(****************************************************************************************************<br>
© Syntegon Group.<br>
All rights reserved, also regarding any disposal, exploitation, reproduction, editing, distribution,<br>
as well as in the event of applications for industrial property rights.<br>
*****************************************************************************************************<br>
DESCRIPTION:<br>
Passes the effective pose, origin shift and zones on to the component's Syn_Visu FB; for m_PassOn of the<br>
derived FB, which knows where the visualisation keeps its zone count.<br>
****************************************************************************************************)
METHOD PROTECTED m_PassOnBody : BOOL
VAR_IN_OUT
	vio_Visu							: SynVisu._FB_VisuBodyComponent;	// the component's Syn_Visu FB
END_VAR
VAR_INPUT
	vi_un_VisuZoneCount					: UINT;	// [-] zones the visualisation has now, its stConfig.nZoneCount
END_VAR
m_PassOnBody := TRUE;
vio_Visu.m_SetPose(vi_Pose := vo_Config.stActive.stPose);
vio_Visu.m_SetOriginShift(vi_lr_X := vo_Config.stActive.stOriginShift.fX, vi_lr_Y := vo_Config.stActive.stOriginShift.fY,
	vi_lr_Z := vo_Config.stActive.stOriginShift.fZ);
m_PassOnZones(vio_Visu := vio_Visu, vio_aZones := vo_Config.stActive.aZones, vi_un_Count := vo_Config.stActive.nZoneCount,
	vi_un_VisuCount := vi_un_VisuZoneCount);
END_METHOD

(****************************************************************************************************<br>
© Syntegon Group.<br>
All rights reserved, also regarding any disposal, exploitation, reproduction, editing, distribution,<br>
as well as in the event of applications for industrial property rights.<br>
*****************************************************************************************************<br>
DESCRIPTION:<br>
Effective pose (MCS), for the application's logic.<br>
****************************************************************************************************)
METHOD m_Pose : SynVisu.ST_VisuPose
m_Pose := vo_Config.stActive.stPose;
END_METHOD

END_FUNCTION_BLOCK

// ---- POUs/_FB_ConfigCartesian.TcPOU
(****************************************************************************************************<br>
© Syntegon Group.<br>
All rights reserved, also regarding any disposal, exploitation, reproduction, editing, distribution,<br>
as well as in the event of applications for industrial property rights.<br>
*****************************************************************************************************<br>
DESCRIPTION:<br>
Parameter set of one Cartesian robot (ADR 0017): its pose, origin shift, zones, gripper fingers, limit area and<br>
TCP limit area, written by the configurator, taken over when the application allows it.<br>
Typical cycle:<br>
  fb_CartParam.m_Register(vio_Manifest := GVL_Config.stManifest, vi_udn_Id := fb_Cart.m_Id());<br>
  fb_CartParam.m_Cycle(vio_Default := CartDefault, vio_Set := CartSet, vi_b_ApplyAllowed := b_Stopped);<br>
  fb_Cart.m_Configure(vi_lr_XMin := 0, ...);<br>
  fb_CartParam.m_PassOn(vio_Visu := fb_Cart);<br>
The application's logic takes its zones and limit areas from m_Active, not from its own constants.<br>
*****************************************************************************************************<br>
OUTPUT VALUES:<br>
vo_Config is the contract structure the gateway reads and writes at the path in the config manifest.<br>
*****************************************************************************************************<br>
VERSION         ¦ DATE       ¦ NAME      ¦ CHANGE<br>
Syn_Config 1.1.0 ¦ 2026-11-10 ¦ J.Willner ¦ New<br>
Syn_Config 2.0.0 ¦ 2026-11-11 ¦ J.Willner ¦ Gripper fingers with their offsets, m_Invalid (ADR 0018)<br>
Syn_Config 2.3.0 ¦ 2026-11-14 ¦ J.Willner ¦ m_Cycle through m_HandleStaging; m_PassOn passes the pose on<br>
****************************************************************************************************)
FUNCTION_BLOCK _FB_ConfigCartesian EXTENDS _FB_ConfigComponent
VAR_OUTPUT
	vo_Config							: ST_ConfigCartesian;	// contract structure of the gateway
END_VAR

(****************************************************************************************************<br>
© Syntegon Group.<br>
All rights reserved, also regarding any disposal, exploitation, reproduction, editing, distribution,<br>
as well as in the event of applications for industrial property rights.<br>
*****************************************************************************************************<br>
DESCRIPTION:<br>
All effective values (zones, limit areas, ...), for the application's own logic.<br>
****************************************************************************************************)
METHOD m_Active : ST_ConfigCartesianParam
m_Active := vo_Config.stActive;
END_METHOD

(****************************************************************************************************<br>
© Syntegon Group.<br>
All rights reserved, also regarding any disposal, exploitation, reproduction, editing, distribution,<br>
as well as in the event of applications for industrial property rights.<br>
*****************************************************************************************************<br>
DESCRIPTION:<br>
A Cartesian robot.<br>
****************************************************************************************************)
METHOD PROTECTED m_ComponentType : SynVisu.E_VisuComponentType
m_ComponentType := SynVisu.E_VisuComponentType.CARTESIAN;
END_METHOD

(****************************************************************************************************<br>
© Syntegon Group.<br>
All rights reserved, also regarding any disposal, exploitation, reproduction, editing, distribution,<br>
as well as in the event of applications for industrial property rights.<br>
*****************************************************************************************************<br>
DESCRIPTION:<br>
Every cycle: handles a staged set or a reset (a set only while vi_b_ApplyAllowed), keeps the active set in<br>
vio_Set and gives the effective values in vo_Config.stActive: the active set while one is valid, else the<br>
program values vio_Default.<br>
*****************************************************************************************************<br>
OUTPUT VALUES:<br>
TRUE in the cycle a set was taken over or reset.<br>
****************************************************************************************************)
METHOD m_Cycle : BOOL
VAR_IN_OUT CONSTANT
	vio_Default							: ST_ConfigCartesianParam;	// the application's program values
END_VAR
VAR_IN_OUT
	vio_Set								: ST_ConfigCartesianSet;	// the application's VAR PERSISTENT active set
END_VAR
VAR_INPUT
	vi_b_ApplyAllowed					: BOOL;	// [-] a staged set may be taken over now, e.g. while the machine stands
END_VAR
VAR
	b_TempTakeOver						: BOOL;	// the staged set was taken over: copy it
END_VAR
m_Cycle := m_HandleStaging(vio_Staging := vo_Config.stStaging, vio_Status := vo_Config.stStatus, vio_b_Valid := vio_Set.bValid,
	vio_udn_Version := vio_Set.nVersion, vio_udn_LastVersion := vio_Set.nLastVersion, vi_b_ApplyAllowed := vi_b_ApplyAllowed,
	vo_b_TakeOver => b_TempTakeOver);
IF b_TempTakeOver THEN
	vio_Set.stParam := vo_Config.stStaged;
END_IF


(****************************************************************************************************
EFFECTIVE VALUES
****************************************************************************************************)
IF vio_Set.bValid THEN
	vo_Config.stActive := vio_Set.stParam;
ELSE
	vo_Config.stActive := vio_Default;
END_IF
END_METHOD

(****************************************************************************************************<br>
© Syntegon Group.<br>
All rights reserved, also regarding any disposal, exploitation, reproduction, editing, distribution,<br>
as well as in the event of applications for industrial property rights.<br>
*****************************************************************************************************<br>
DESCRIPTION:<br>
Why a staged set cannot be taken over; '' when it can: more zones or fingers than the lists hold, a zone on no<br>
conveyor (id 0), or a finger without a diameter or height.<br>
****************************************************************************************************)
METHOD PROTECTED m_InvalidStaged : STRING(80)
m_InvalidStaged := m_InvalidZones(vio_aZones := vo_Config.stStaged.aZones, vi_un_Count := vo_Config.stStaged.nZoneCount);
IF m_InvalidStaged = '' THEN
	m_InvalidStaged := m_InvalidFingers(vio_aFingers := vo_Config.stStaged.aFingers, vi_un_Count := vo_Config.stStaged.nFingerCount);
END_IF
END_METHOD

(****************************************************************************************************<br>
© Syntegon Group.<br>
All rights reserved, also regarding any disposal, exploitation, reproduction, editing, distribution,<br>
as well as in the event of applications for industrial property rights.<br>
*****************************************************************************************************<br>
DESCRIPTION:<br>
Passes the effective pose, origin shift, limit areas, zones and fingers on to the robot's Syn_Visu FB, so the<br>
visualisation shows what the machine uses; the strokes and rail height (hardware) stay with the application's<br>
m_Configure call. Call it after m_Cycle, every cycle; Syn_Visu's config version only changes when a value does.<br>
****************************************************************************************************)
METHOD m_PassOn : BOOL
VAR_IN_OUT
	vio_Visu							: SynVisu._FB_VisuCartesian;	// the robot's Syn_Visu FB
END_VAR
m_PassOn := TRUE;
vio_Visu.m_SetPose(vi_Pose := vo_Config.stActive.stPose);
vio_Visu.m_SetOriginShift(vi_lr_X := vo_Config.stActive.stOriginShift.fX, vi_lr_Y := vo_Config.stActive.stOriginShift.fY,
	vi_lr_Z := vo_Config.stActive.stOriginShift.fZ);
m_PassOnLimitAreas(vio_Visu := vio_Visu, vio_LimitArea := vo_Config.stActive.stLimitArea,
	vio_TcpLimitArea := vo_Config.stActive.stTcpLimitArea);
m_PassOnZones(vio_Visu := vio_Visu, vio_aZones := vo_Config.stActive.aZones, vi_un_Count := vo_Config.stActive.nZoneCount,
	vi_un_VisuCount := vio_Visu.vo_Visu.stConfig.nZoneCount);
m_PassOnFingers(vio_Visu := vio_Visu, vio_aFingers := vo_Config.stActive.aFingers,
	vi_un_Count := vo_Config.stActive.nFingerCount, vi_un_VisuCount := vio_Visu.vo_Visu.stConfig.nFingerCount);
END_METHOD

(****************************************************************************************************<br>
© Syntegon Group.<br>
All rights reserved, also regarding any disposal, exploitation, reproduction, editing, distribution,<br>
as well as in the event of applications for industrial property rights.<br>
*****************************************************************************************************<br>
DESCRIPTION:<br>
Effective pose of the axis origin (MCS), for the application's logic.<br>
****************************************************************************************************)
METHOD m_Pose : SynVisu.ST_VisuPose
m_Pose := vo_Config.stActive.stPose;
END_METHOD

END_FUNCTION_BLOCK

// ---- POUs/_FB_ConfigConveyor.TcPOU
(****************************************************************************************************<br>
© Syntegon Group.<br>
All rights reserved, also regarding any disposal, exploitation, reproduction, editing, distribution,<br>
as well as in the event of applications for industrial property rights.<br>
*****************************************************************************************************<br>
DESCRIPTION:<br>
Parameter set of one conveyor (ADR 0017): its pose, origin shift and product types, written by the configurator,<br>
taken over when the application allows it. Typical cycle, before the Syn_Visu calls of the conveyor:<br>
  fb_InfeedParam.m_Register(vio_Manifest := GVL_Config.stManifest, vi_udn_Id := fb_Infeed.m_Id());<br>
  fb_InfeedParam.m_Cycle(vio_Default := InfeedDefault, vio_Set := InfeedSet, vi_b_ApplyAllowed := b_Stopped);<br>
  fb_Infeed.m_Configure(vi_lr_Length := 3000, vi_lr_Width := 400);<br>
  fb_InfeedParam.m_PassOn(vio_Visu := fb_Infeed);<br>
InfeedSet is the application's VAR PERSISTENT ST_ConfigConveyorSet; InfeedDefault its program values.<br>
*****************************************************************************************************<br>
OUTPUT VALUES:<br>
vo_Config is the contract structure the gateway reads and writes at the path in the config manifest.<br>
*****************************************************************************************************<br>
VERSION         ¦ DATE       ¦ NAME      ¦ CHANGE<br>
Syn_Config 1.0.0 ¦ 2026-11-10 ¦ J.Willner ¦ First version<br>
Syn_Config 2.3.0 ¦ 2026-11-14 ¦ J.Willner ¦ m_Cycle through m_HandleStaging; m_PassOn passes the pose on<br>
****************************************************************************************************)
FUNCTION_BLOCK _FB_ConfigConveyor EXTENDS _FB_ConfigComponent
VAR_OUTPUT
	vo_Config							: ST_ConfigConveyor;	// contract structure of the gateway
END_VAR

(****************************************************************************************************<br>
© Syntegon Group.<br>
All rights reserved, also regarding any disposal, exploitation, reproduction, editing, distribution,<br>
as well as in the event of applications for industrial property rights.<br>
*****************************************************************************************************<br>
DESCRIPTION:<br>
All effective values (origin shift, product types, ...), for the application's own logic.<br>
****************************************************************************************************)
METHOD m_Active : ST_ConfigConveyorParam
m_Active := vo_Config.stActive;
END_METHOD

(****************************************************************************************************<br>
© Syntegon Group.<br>
All rights reserved, also regarding any disposal, exploitation, reproduction, editing, distribution,<br>
as well as in the event of applications for industrial property rights.<br>
*****************************************************************************************************<br>
DESCRIPTION:<br>
A conveyor.<br>
****************************************************************************************************)
METHOD PROTECTED m_ComponentType : SynVisu.E_VisuComponentType
m_ComponentType := SynVisu.E_VisuComponentType.CONVEYOR;
END_METHOD

(****************************************************************************************************<br>
© Syntegon Group.<br>
All rights reserved, also regarding any disposal, exploitation, reproduction, editing, distribution,<br>
as well as in the event of applications for industrial property rights.<br>
*****************************************************************************************************<br>
DESCRIPTION:<br>
Every cycle: handles a staged set or a reset (a set only while vi_b_ApplyAllowed), keeps the active set in<br>
vio_Set and gives the effective values in vo_Config.stActive: the active set while one is valid, else the<br>
program values vio_Default.<br>
*****************************************************************************************************<br>
OUTPUT VALUES:<br>
TRUE in the cycle a set was taken over or reset.<br>
****************************************************************************************************)
METHOD m_Cycle : BOOL
VAR_IN_OUT CONSTANT
	vio_Default							: ST_ConfigConveyorParam;	// the application's program values
END_VAR
VAR_IN_OUT
	vio_Set								: ST_ConfigConveyorSet;	// the application's VAR PERSISTENT active set
END_VAR
VAR_INPUT
	vi_b_ApplyAllowed					: BOOL;	// [-] a staged set may be taken over now, e.g. while the machine stands
END_VAR
VAR
	b_TempTakeOver						: BOOL;	// the staged set was taken over: copy it
END_VAR
m_Cycle := m_HandleStaging(vio_Staging := vo_Config.stStaging, vio_Status := vo_Config.stStatus, vio_b_Valid := vio_Set.bValid,
	vio_udn_Version := vio_Set.nVersion, vio_udn_LastVersion := vio_Set.nLastVersion, vi_b_ApplyAllowed := vi_b_ApplyAllowed,
	vo_b_TakeOver => b_TempTakeOver);
IF b_TempTakeOver THEN
	vio_Set.stParam := vo_Config.stStaged;
END_IF


(****************************************************************************************************
EFFECTIVE VALUES
****************************************************************************************************)
IF vio_Set.bValid THEN
	vo_Config.stActive := vio_Set.stParam;
ELSE
	vo_Config.stActive := vio_Default;
END_IF
END_METHOD

(****************************************************************************************************<br>
© Syntegon Group.<br>
All rights reserved, also regarding any disposal, exploitation, reproduction, editing, distribution,<br>
as well as in the event of applications for industrial property rights.<br>
*****************************************************************************************************<br>
DESCRIPTION:<br>
Why a staged set cannot be taken over; '' when it can: more product types than the list holds, a product type<br>
without a number or a number used twice.<br>
****************************************************************************************************)
METHOD PROTECTED m_InvalidStaged : STRING(80)
VAR
	un_TempIndex						: UINT;
	un_TempOther						: UINT;
END_VAR
m_InvalidStaged := '';
IF vo_Config.stStaged.nProductTypeCount > SynVisu.VISU_GlobalConst_Param.VISU_un_MAX_PRODUCT_TYPES THEN
	m_InvalidStaged := CONCAT('More than ', CONCAT(UINT_TO_STRING(SynVisu.VISU_GlobalConst_Param.VISU_un_MAX_PRODUCT_TYPES), ' product types'));
	RETURN;
END_IF
un_TempIndex := 0;
WHILE un_TempIndex < vo_Config.stStaged.nProductTypeCount DO
	IF vo_Config.stStaged.aProductTypes[un_TempIndex].nId = 0 THEN
		m_InvalidStaged := 'A product type without a number';
		RETURN;
	END_IF
	un_TempOther := 0;
	WHILE un_TempOther < un_TempIndex DO
		IF vo_Config.stStaged.aProductTypes[un_TempOther].nId = vo_Config.stStaged.aProductTypes[un_TempIndex].nId THEN
			m_InvalidStaged := CONCAT('Product type ',
				CONCAT(UDINT_TO_STRING(vo_Config.stStaged.aProductTypes[un_TempIndex].nId), ' is defined twice'));
			RETURN;
		END_IF
		un_TempOther := un_TempOther + 1;
	END_WHILE
	un_TempIndex := un_TempIndex + 1;
END_WHILE
END_METHOD

(****************************************************************************************************<br>
© Syntegon Group.<br>
All rights reserved, also regarding any disposal, exploitation, reproduction, editing, distribution,<br>
as well as in the event of applications for industrial property rights.<br>
*****************************************************************************************************<br>
DESCRIPTION:<br>
Passes the effective pose, origin shift and product types on to the conveyor's Syn_Visu FB, so the<br>
visualisation shows what the machine uses; the belt's length and width (hardware) stay with the application's<br>
m_Configure call. Call it after m_Cycle, every cycle; Syn_Visu's config version only changes when a value does.<br>
*****************************************************************************************************<br>
LIMITS:<br>
Syn_Visu cannot remove a product type: one the set no longer has stays in the visualisation until the<br>
application restarts (the configurator warns of the difference).<br>
****************************************************************************************************)
METHOD m_PassOn : BOOL
VAR_IN_OUT
	vio_Visu							: SynVisu._FB_VisuConveyor;	// the conveyor's Syn_Visu FB
END_VAR
VAR
	un_TempIndex						: UINT;
END_VAR
m_PassOn := TRUE;
vio_Visu.m_SetPose(vi_Pose := vo_Config.stActive.stPose);
vio_Visu.m_SetOriginShift(vi_lr_X := vo_Config.stActive.stOriginShift.fX, vi_lr_Y := vo_Config.stActive.stOriginShift.fY,
	vi_lr_Z := vo_Config.stActive.stOriginShift.fZ);
un_TempIndex := 0;
WHILE un_TempIndex < vo_Config.stActive.nProductTypeCount
	AND un_TempIndex < SynVisu.VISU_GlobalConst_Param.VISU_un_MAX_PRODUCT_TYPES
DO
	vio_Visu.m_SetProductType(vi_udn_Id := vo_Config.stActive.aProductTypes[un_TempIndex].nId,
		vi_lr_Length := vo_Config.stActive.aProductTypes[un_TempIndex].fLength,
		vi_lr_Width := vo_Config.stActive.aProductTypes[un_TempIndex].fWidth,
		vi_lr_Height := vo_Config.stActive.aProductTypes[un_TempIndex].fHeight,
		vi_e_Shape := vo_Config.stActive.aProductTypes[un_TempIndex].eShape,
		vi_lr_CornerRadius := vo_Config.stActive.aProductTypes[un_TempIndex].fCornerRadius);
	un_TempIndex := un_TempIndex + 1;
END_WHILE
END_METHOD

(****************************************************************************************************<br>
© Syntegon Group.<br>
All rights reserved, also regarding any disposal, exploitation, reproduction, editing, distribution,<br>
as well as in the event of applications for industrial property rights.<br>
*****************************************************************************************************<br>
DESCRIPTION:<br>
Effective pose of the belt start (MCS), for the application's logic.<br>
****************************************************************************************************)
METHOD m_Pose : SynVisu.ST_VisuPose
m_Pose := vo_Config.stActive.stPose;
END_METHOD

END_FUNCTION_BLOCK

// ---- POUs/_FB_ConfigDelta.TcPOU
(****************************************************************************************************<br>
© Syntegon Group.<br>
All rights reserved, also regarding any disposal, exploitation, reproduction, editing, distribution,<br>
as well as in the event of applications for industrial property rights.<br>
*****************************************************************************************************<br>
DESCRIPTION:<br>
Parameter set of one Delta robot (ADR 0017): its pose, origin shift, zones, gripper fingers, working area,<br>
limit area and TCP limit area, written by the configurator, taken over when the application allows it.<br>
Typical cycle:<br>
  fb_Delta1Param.m_Register(vio_Manifest := GVL_Config.stManifest, vi_udn_Id := fb_Delta1.m_Id());<br>
  fb_Delta1Param.m_Cycle(vio_Default := Delta1Default, vio_Set := Delta1Set, vi_b_ApplyAllowed := b_Stopped);<br>
  fb_Delta1.m_Configure(vi_lr_BaseRadius := 200, ...);<br>
  fb_Delta1Param.m_PassOn(vio_Visu := fb_Delta1);<br>
The application's pick logic takes its zones from m_Zone / m_Active, not from its own constants.<br>
*****************************************************************************************************<br>
OUTPUT VALUES:<br>
vo_Config is the contract structure the gateway reads and writes at the path in the config manifest.<br>
*****************************************************************************************************<br>
VERSION         ¦ DATE       ¦ NAME      ¦ CHANGE<br>
Syn_Config 1.0.0 ¦ 2026-11-10 ¦ J.Willner ¦ First version<br>
Syn_Config 1.1.0 ¦ 2026-11-10 ¦ J.Willner ¦ m_PassOn, m_Invalid through the shared helpers<br>
Syn_Config 2.0.0 ¦ 2026-11-11 ¦ J.Willner ¦ Gripper fingers with their offsets (ADR 0018)<br>
Syn_Config 2.3.0 ¦ 2026-11-14 ¦ J.Willner ¦ m_Cycle through m_HandleStaging; m_PassOn passes the pose on<br>
****************************************************************************************************)
FUNCTION_BLOCK _FB_ConfigDelta EXTENDS _FB_ConfigComponent
VAR_OUTPUT
	vo_Config							: ST_ConfigDelta;	// contract structure of the gateway
END_VAR

(****************************************************************************************************<br>
© Syntegon Group.<br>
All rights reserved, also regarding any disposal, exploitation, reproduction, editing, distribution,<br>
as well as in the event of applications for industrial property rights.<br>
*****************************************************************************************************<br>
DESCRIPTION:<br>
All effective values (zones, working and limit areas, ...), for the application's own logic.<br>
****************************************************************************************************)
METHOD m_Active : ST_ConfigDeltaParam
m_Active := vo_Config.stActive;
END_METHOD

(****************************************************************************************************<br>
© Syntegon Group.<br>
All rights reserved, also regarding any disposal, exploitation, reproduction, editing, distribution,<br>
as well as in the event of applications for industrial property rights.<br>
*****************************************************************************************************<br>
DESCRIPTION:<br>
A Delta robot.<br>
****************************************************************************************************)
METHOD PROTECTED m_ComponentType : SynVisu.E_VisuComponentType
m_ComponentType := SynVisu.E_VisuComponentType.DELTA;
END_METHOD

(****************************************************************************************************<br>
© Syntegon Group.<br>
All rights reserved, also regarding any disposal, exploitation, reproduction, editing, distribution,<br>
as well as in the event of applications for industrial property rights.<br>
*****************************************************************************************************<br>
DESCRIPTION:<br>
Every cycle: handles a staged set or a reset (a set only while vi_b_ApplyAllowed), keeps the active set in<br>
vio_Set and gives the effective values in vo_Config.stActive: the active set while one is valid, else the<br>
program values vio_Default.<br>
*****************************************************************************************************<br>
OUTPUT VALUES:<br>
TRUE in the cycle a set was taken over or reset.<br>
****************************************************************************************************)
METHOD m_Cycle : BOOL
VAR_IN_OUT CONSTANT
	vio_Default							: ST_ConfigDeltaParam;	// the application's program values
END_VAR
VAR_IN_OUT
	vio_Set								: ST_ConfigDeltaSet;	// the application's VAR PERSISTENT active set
END_VAR
VAR_INPUT
	vi_b_ApplyAllowed					: BOOL;	// [-] a staged set may be taken over now, e.g. while the machine stands
END_VAR
VAR
	b_TempTakeOver						: BOOL;	// the staged set was taken over: copy it
END_VAR
m_Cycle := m_HandleStaging(vio_Staging := vo_Config.stStaging, vio_Status := vo_Config.stStatus, vio_b_Valid := vio_Set.bValid,
	vio_udn_Version := vio_Set.nVersion, vio_udn_LastVersion := vio_Set.nLastVersion, vi_b_ApplyAllowed := vi_b_ApplyAllowed,
	vo_b_TakeOver => b_TempTakeOver);
IF b_TempTakeOver THEN
	vio_Set.stParam := vo_Config.stStaged;
END_IF


(****************************************************************************************************
EFFECTIVE VALUES
****************************************************************************************************)
IF vio_Set.bValid THEN
	vo_Config.stActive := vio_Set.stParam;
ELSE
	vo_Config.stActive := vio_Default;
END_IF
END_METHOD

(****************************************************************************************************<br>
© Syntegon Group.<br>
All rights reserved, also regarding any disposal, exploitation, reproduction, editing, distribution,<br>
as well as in the event of applications for industrial property rights.<br>
*****************************************************************************************************<br>
DESCRIPTION:<br>
Why a staged set cannot be taken over; '' when it can: more zones or fingers than the lists hold, a zone on no<br>
conveyor (id 0), or a finger without a diameter or height.<br>
****************************************************************************************************)
METHOD PROTECTED m_InvalidStaged : STRING(80)
m_InvalidStaged := m_InvalidZones(vio_aZones := vo_Config.stStaged.aZones, vi_un_Count := vo_Config.stStaged.nZoneCount);
IF m_InvalidStaged = '' THEN
	m_InvalidStaged := m_InvalidFingers(vio_aFingers := vo_Config.stStaged.aFingers, vi_un_Count := vo_Config.stStaged.nFingerCount);
END_IF
END_METHOD

(****************************************************************************************************<br>
© Syntegon Group.<br>
All rights reserved, also regarding any disposal, exploitation, reproduction, editing, distribution,<br>
as well as in the event of applications for industrial property rights.<br>
*****************************************************************************************************<br>
DESCRIPTION:<br>
Passes the effective pose, origin shift, working area, limit areas, zones and fingers on to the Delta's<br>
Syn_Visu FB, so the visualisation shows what the machine uses; the arm geometry (hardware) stays with the<br>
application's m_Configure call. Call it after m_Cycle, every cycle; Syn_Visu's config version only changes when a<br>
value does (zones and fingers are cleared only when the set has fewer than the visualisation).<br>
****************************************************************************************************)
METHOD m_PassOn : BOOL
VAR_IN_OUT
	vio_Visu							: SynVisu._FB_VisuDelta;	// the Delta's Syn_Visu FB
END_VAR
m_PassOn := TRUE;
vio_Visu.m_SetPose(vi_Pose := vo_Config.stActive.stPose);
vio_Visu.m_SetOriginShift(vi_lr_X := vo_Config.stActive.stOriginShift.fX, vi_lr_Y := vo_Config.stActive.stOriginShift.fY,
	vi_lr_Z := vo_Config.stActive.stOriginShift.fZ);
vio_Visu.m_SetWorkingArea(vi_lr_Radius := vo_Config.stActive.stWorkingArea.fRadius,
	vi_lr_ZMin := vo_Config.stActive.stWorkingArea.fZMin, vi_lr_ZMax := vo_Config.stActive.stWorkingArea.fZMax,
	vi_lr_ConeHeight := vo_Config.stActive.stWorkingArea.fConeHeight,
	vi_lr_ConeBottomRadius := vo_Config.stActive.stWorkingArea.fConeBottomRadius);
m_PassOnLimitAreas(vio_Visu := vio_Visu, vio_LimitArea := vo_Config.stActive.stLimitArea,
	vio_TcpLimitArea := vo_Config.stActive.stTcpLimitArea);
m_PassOnZones(vio_Visu := vio_Visu, vio_aZones := vo_Config.stActive.aZones, vi_un_Count := vo_Config.stActive.nZoneCount,
	vi_un_VisuCount := vio_Visu.vo_Visu.stConfig.nZoneCount);
m_PassOnFingers(vio_Visu := vio_Visu, vio_aFingers := vo_Config.stActive.aFingers,
	vi_un_Count := vo_Config.stActive.nFingerCount, vi_un_VisuCount := vio_Visu.vo_Visu.stConfig.nFingerCount);
END_METHOD

(****************************************************************************************************<br>
© Syntegon Group.<br>
All rights reserved, also regarding any disposal, exploitation, reproduction, editing, distribution,<br>
as well as in the event of applications for industrial property rights.<br>
*****************************************************************************************************<br>
DESCRIPTION:<br>
Effective pose of the base centre (MCS), for the application's logic.<br>
****************************************************************************************************)
METHOD m_Pose : SynVisu.ST_VisuPose
m_Pose := vo_Config.stActive.stPose;
END_METHOD

(****************************************************************************************************<br>
© Syntegon Group.<br>
All rights reserved, also regarding any disposal, exploitation, reproduction, editing, distribution,<br>
as well as in the event of applications for industrial property rights.<br>
*****************************************************************************************************<br>
DESCRIPTION:<br>
Effective zone vi_un_Zone (1-based, as in Syn_Visu's m_SetZone), for the application's pick and place logic.<br>
*****************************************************************************************************<br>
OUTPUT VALUES:<br>
A zone with nConveyorId = 0 for a number outside 1..m_ZoneCount().<br>
****************************************************************************************************)
METHOD m_Zone : SynVisu.ST_VisuZone
VAR_INPUT
	vi_un_Zone							: UINT;	// [-] 1-based
END_VAR
IF vi_un_Zone >= 1 AND vi_un_Zone <= vo_Config.stActive.nZoneCount
	AND vi_un_Zone <= SynVisu.VISU_GlobalConst_Param.VISU_un_MAX_ZONES
THEN
	m_Zone := vo_Config.stActive.aZones[vi_un_Zone - 1];
END_IF
END_METHOD

(****************************************************************************************************<br>
© Syntegon Group.<br>
All rights reserved, also regarding any disposal, exploitation, reproduction, editing, distribution,<br>
as well as in the event of applications for industrial property rights.<br>
*****************************************************************************************************<br>
DESCRIPTION:<br>
Number of effective zones.<br>
****************************************************************************************************)
METHOD m_ZoneCount : UINT
m_ZoneCount := vo_Config.stActive.nZoneCount;
END_METHOD

END_FUNCTION_BLOCK

// ---- POUs/_FB_ConfigSensor.TcPOU
(****************************************************************************************************<br>
© Syntegon Group.<br>
All rights reserved, also regarding any disposal, exploitation, reproduction, editing, distribution,<br>
as well as in the event of applications for industrial property rights.<br>
*****************************************************************************************************<br>
DESCRIPTION:<br>
Parameter set of one product sensor (ADR 0017): its pose, origin shift and zones. See _FB_ConfigBodyComponent.<br>
*****************************************************************************************************<br>
VERSION         ¦ DATE       ¦ NAME      ¦ CHANGE<br>
Syn_Config 1.1.0 ¦ 2026-11-10 ¦ J.Willner ¦ New<br>
Syn_Config 2.3.0 ¦ 2026-11-14 ¦ J.Willner ¦ m_PassOn passes the pose on<br>
****************************************************************************************************)
FUNCTION_BLOCK _FB_ConfigSensor EXTENDS _FB_ConfigBodyComponent

(****************************************************************************************************<br>
© Syntegon Group.<br>
All rights reserved, also regarding any disposal, exploitation, reproduction, editing, distribution,<br>
as well as in the event of applications for industrial property rights.<br>
*****************************************************************************************************<br>
DESCRIPTION:<br>
A product sensor.<br>
****************************************************************************************************)
METHOD PROTECTED m_ComponentType : SynVisu.E_VisuComponentType
m_ComponentType := SynVisu.E_VisuComponentType.SENSOR;
END_METHOD

(****************************************************************************************************<br>
© Syntegon Group.<br>
All rights reserved, also regarding any disposal, exploitation, reproduction, editing, distribution,<br>
as well as in the event of applications for industrial property rights.<br>
*****************************************************************************************************<br>
DESCRIPTION:<br>
Passes the effective pose, origin shift and zones on to the sensor's Syn_Visu FB; the beam length (hardware)<br>
stays with the application's m_Configure call. Call it after m_Cycle, every cycle.<br>
****************************************************************************************************)
METHOD m_PassOn : BOOL
VAR_IN_OUT
	vio_Visu							: SynVisu._FB_VisuSensor;	// the sensor's Syn_Visu FB
END_VAR
m_PassOn := m_PassOnBody(vio_Visu := vio_Visu, vi_un_VisuZoneCount := vio_Visu.vo_Visu.stConfig.nZoneCount);
END_METHOD

END_FUNCTION_BLOCK

// ---- POUs/_FB_ConfigStation.TcPOU
(****************************************************************************************************<br>
© Syntegon Group.<br>
All rights reserved, also regarding any disposal, exploitation, reproduction, editing, distribution,<br>
as well as in the event of applications for industrial property rights.<br>
*****************************************************************************************************<br>
DESCRIPTION:<br>
Parameter set of one station (reject unit, labeller, ..., ADR 0017): its pose, origin shift and zones. See<br>
_FB_ConfigBodyComponent.<br>
*****************************************************************************************************<br>
VERSION         ¦ DATE       ¦ NAME      ¦ CHANGE<br>
Syn_Config 1.1.0 ¦ 2026-11-10 ¦ J.Willner ¦ New<br>
Syn_Config 2.3.0 ¦ 2026-11-14 ¦ J.Willner ¦ m_PassOn passes the pose on<br>
****************************************************************************************************)
FUNCTION_BLOCK _FB_ConfigStation EXTENDS _FB_ConfigBodyComponent

(****************************************************************************************************<br>
© Syntegon Group.<br>
All rights reserved, also regarding any disposal, exploitation, reproduction, editing, distribution,<br>
as well as in the event of applications for industrial property rights.<br>
*****************************************************************************************************<br>
DESCRIPTION:<br>
A station.<br>
****************************************************************************************************)
METHOD PROTECTED m_ComponentType : SynVisu.E_VisuComponentType
m_ComponentType := SynVisu.E_VisuComponentType.STATION;
END_METHOD

(****************************************************************************************************<br>
© Syntegon Group.<br>
All rights reserved, also regarding any disposal, exploitation, reproduction, editing, distribution,<br>
as well as in the event of applications for industrial property rights.<br>
*****************************************************************************************************<br>
DESCRIPTION:<br>
Passes the effective pose, origin shift and zones on to the station's Syn_Visu FB; its bodies stay the<br>
application's (hardware). Call it after m_Cycle, every cycle.<br>
****************************************************************************************************)
METHOD m_PassOn : BOOL
VAR_IN_OUT
	vio_Visu							: SynVisu._FB_VisuStation;	// the station's Syn_Visu FB
END_VAR
m_PassOn := m_PassOnBody(vio_Visu := vio_Visu, vi_un_VisuZoneCount := vio_Visu.vo_Visu.stConfig.nZoneCount);
END_METHOD

END_FUNCTION_BLOCK

// ---- POUs/_FB_ConfigVision.TcPOU
(****************************************************************************************************<br>
© Syntegon Group.<br>
All rights reserved, also regarding any disposal, exploitation, reproduction, editing, distribution,<br>
as well as in the event of applications for industrial property rights.<br>
*****************************************************************************************************<br>
DESCRIPTION:<br>
Parameter set of one vision system (ADR 0017): its pose, origin shift and zones. See _FB_ConfigBodyComponent.<br>
*****************************************************************************************************<br>
VERSION         ¦ DATE       ¦ NAME      ¦ CHANGE<br>
Syn_Config 1.1.0 ¦ 2026-11-10 ¦ J.Willner ¦ New<br>
Syn_Config 2.3.0 ¦ 2026-11-14 ¦ J.Willner ¦ m_PassOn passes the pose on<br>
****************************************************************************************************)
FUNCTION_BLOCK _FB_ConfigVision EXTENDS _FB_ConfigBodyComponent

(****************************************************************************************************<br>
© Syntegon Group.<br>
All rights reserved, also regarding any disposal, exploitation, reproduction, editing, distribution,<br>
as well as in the event of applications for industrial property rights.<br>
*****************************************************************************************************<br>
DESCRIPTION:<br>
A vision system.<br>
****************************************************************************************************)
METHOD PROTECTED m_ComponentType : SynVisu.E_VisuComponentType
m_ComponentType := SynVisu.E_VisuComponentType.VISION;
END_METHOD

(****************************************************************************************************<br>
© Syntegon Group.<br>
All rights reserved, also regarding any disposal, exploitation, reproduction, editing, distribution,<br>
as well as in the event of applications for industrial property rights.<br>
*****************************************************************************************************<br>
DESCRIPTION:<br>
Passes the effective pose, origin shift and zones on to the vision system's Syn_Visu FB; the field of view<br>
(hardware) stays with the application's m_Configure call. Call it after m_Cycle, every cycle.<br>
****************************************************************************************************)
METHOD m_PassOn : BOOL
VAR_IN_OUT
	vio_Visu							: SynVisu._FB_VisuVision;	// the vision system's Syn_Visu FB
END_VAR
m_PassOn := m_PassOnBody(vio_Visu := vio_Visu, vi_un_VisuZoneCount := vio_Visu.vo_Visu.stConfig.nZoneCount);
END_METHOD

END_FUNCTION_BLOCK

// ---- POUs/_FB_ConfigXtsGantry.TcPOU
(****************************************************************************************************<br>
© Syntegon Group.<br>
All rights reserved, also regarding any disposal, exploitation, reproduction, editing, distribution,<br>
as well as in the event of applications for industrial property rights.<br>
*****************************************************************************************************<br>
DESCRIPTION:<br>
Parameter set of one XTS gantry (ADR 0017): its pose, origin shift, track modules, zones, gripper fingers,<br>
limit area and TCP limit area, written by the configurator, taken over when the application allows it.<br>
Typical cycle:<br>
  fb_IdhParam.m_Register(vio_Manifest := GVL_Config.stManifest, vi_udn_Id := fb_Idh.m_Id());<br>
  fb_IdhParam.m_Cycle(vio_Default := IdhDefault, vio_Set := IdhSet, vi_b_ApplyAllowed := b_Stopped);<br>
  fb_Idh.m_Configure(vi_lr_XMin := 0, ...);<br>
  fb_IdhParam.m_PassOn(vio_Visu := fb_Idh);<br>
The application's logic takes its track and zones from m_Active, not from its own constants.<br>
*****************************************************************************************************<br>
OUTPUT VALUES:<br>
vo_Config is the contract structure the gateway reads and writes at the path in the config manifest.<br>
*****************************************************************************************************<br>
VERSION         ¦ DATE       ¦ NAME      ¦ CHANGE<br>
Syn_Config 1.1.0 ¦ 2026-11-10 ¦ J.Willner ¦ New<br>
Syn_Config 2.0.0 ¦ 2026-11-11 ¦ J.Willner ¦ Gripper fingers with their offsets (ADR 0018)<br>
Syn_Config 2.3.0 ¦ 2026-11-14 ¦ J.Willner ¦ m_Cycle through m_HandleStaging; m_PassOn passes the pose on<br>
****************************************************************************************************)
FUNCTION_BLOCK _FB_ConfigXtsGantry EXTENDS _FB_ConfigComponent
VAR_OUTPUT
	vo_Config							: ST_ConfigXtsGantry;	// contract structure of the gateway
END_VAR

(****************************************************************************************************<br>
© Syntegon Group.<br>
All rights reserved, also regarding any disposal, exploitation, reproduction, editing, distribution,<br>
as well as in the event of applications for industrial property rights.<br>
*****************************************************************************************************<br>
DESCRIPTION:<br>
All effective values (track modules, zones, limit areas, ...), for the application's own logic.<br>
****************************************************************************************************)
METHOD m_Active : ST_ConfigXtsGantryParam
m_Active := vo_Config.stActive;
END_METHOD

(****************************************************************************************************<br>
© Syntegon Group.<br>
All rights reserved, also regarding any disposal, exploitation, reproduction, editing, distribution,<br>
as well as in the event of applications for industrial property rights.<br>
*****************************************************************************************************<br>
DESCRIPTION:<br>
An XTS gantry.<br>
****************************************************************************************************)
METHOD PROTECTED m_ComponentType : SynVisu.E_VisuComponentType
m_ComponentType := SynVisu.E_VisuComponentType.XTS_GANTRY;
END_METHOD

(****************************************************************************************************<br>
© Syntegon Group.<br>
All rights reserved, also regarding any disposal, exploitation, reproduction, editing, distribution,<br>
as well as in the event of applications for industrial property rights.<br>
*****************************************************************************************************<br>
DESCRIPTION:<br>
Every cycle: handles a staged set or a reset (a set only while vi_b_ApplyAllowed), keeps the active set in<br>
vio_Set and gives the effective values in vo_Config.stActive: the active set while one is valid, else the<br>
program values vio_Default.<br>
*****************************************************************************************************<br>
OUTPUT VALUES:<br>
TRUE in the cycle a set was taken over or reset.<br>
****************************************************************************************************)
METHOD m_Cycle : BOOL
VAR_IN_OUT CONSTANT
	vio_Default							: ST_ConfigXtsGantryParam;	// the application's program values
END_VAR
VAR_IN_OUT
	vio_Set								: ST_ConfigXtsGantrySet;	// the application's VAR PERSISTENT active set
END_VAR
VAR_INPUT
	vi_b_ApplyAllowed					: BOOL;	// [-] a staged set may be taken over now, e.g. while the machine stands
END_VAR
VAR
	b_TempTakeOver						: BOOL;	// the staged set was taken over: copy it
END_VAR
m_Cycle := m_HandleStaging(vio_Staging := vo_Config.stStaging, vio_Status := vo_Config.stStatus, vio_b_Valid := vio_Set.bValid,
	vio_udn_Version := vio_Set.nVersion, vio_udn_LastVersion := vio_Set.nLastVersion, vi_b_ApplyAllowed := vi_b_ApplyAllowed,
	vo_b_TakeOver => b_TempTakeOver);
IF b_TempTakeOver THEN
	vio_Set.stParam := vo_Config.stStaged;
END_IF


(****************************************************************************************************
EFFECTIVE VALUES
****************************************************************************************************)
IF vio_Set.bValid THEN
	vo_Config.stActive := vio_Set.stParam;
ELSE
	vo_Config.stActive := vio_Default;
END_IF
END_METHOD

(****************************************************************************************************<br>
© Syntegon Group.<br>
All rights reserved, also regarding any disposal, exploitation, reproduction, editing, distribution,<br>
as well as in the event of applications for industrial property rights.<br>
*****************************************************************************************************<br>
DESCRIPTION:<br>
Why a staged set cannot be taken over; '' when it can: a track without modules, more modules, zones or fingers<br>
than the lists hold, a module without a length, a zone on no conveyor (id 0), or a finger without a diameter or<br>
height.<br>
****************************************************************************************************)
METHOD PROTECTED m_InvalidStaged : STRING(80)
m_InvalidStaged := m_InvalidModules(vio_aModules := vo_Config.stStaged.aModules, vi_un_Count := vo_Config.stStaged.nModuleCount);
IF m_InvalidStaged = '' THEN
	m_InvalidStaged := m_InvalidZones(vio_aZones := vo_Config.stStaged.aZones, vi_un_Count := vo_Config.stStaged.nZoneCount);
END_IF
IF m_InvalidStaged = '' THEN
	m_InvalidStaged := m_InvalidFingers(vio_aFingers := vo_Config.stStaged.aFingers, vi_un_Count := vo_Config.stStaged.nFingerCount);
END_IF
END_METHOD

(****************************************************************************************************<br>
© Syntegon Group.<br>
All rights reserved, also regarding any disposal, exploitation, reproduction, editing, distribution,<br>
as well as in the event of applications for industrial property rights.<br>
*****************************************************************************************************<br>
DESCRIPTION:<br>
Passes the effective pose, origin shift, track modules, limit areas, zones and fingers on to the gantry's<br>
Syn_Visu FB, so the visualisation shows what the machine uses; the strokes and tool offsets (hardware) stay with<br>
the application's m_Configure call. Call it after m_Cycle, every cycle; Syn_Visu's config version only changes<br>
when a value does.<br>
****************************************************************************************************)
METHOD m_PassOn : BOOL
VAR_IN_OUT
	vio_Visu							: SynVisu._FB_VisuXtsGantry;	// the gantry's Syn_Visu FB
END_VAR
m_PassOn := TRUE;
vio_Visu.m_SetPose(vi_Pose := vo_Config.stActive.stPose);
vio_Visu.m_SetOriginShift(vi_lr_X := vo_Config.stActive.stOriginShift.fX, vi_lr_Y := vo_Config.stActive.stOriginShift.fY,
	vi_lr_Z := vo_Config.stActive.stOriginShift.fZ);
m_PassOnModules(vio_Visu := vio_Visu, vio_aModules := vo_Config.stActive.aModules,
	vi_un_Count := vo_Config.stActive.nModuleCount, vi_un_VisuCount := vio_Visu.vo_Visu.stConfig.nModuleCount);
m_PassOnLimitAreas(vio_Visu := vio_Visu, vio_LimitArea := vo_Config.stActive.stLimitArea,
	vio_TcpLimitArea := vo_Config.stActive.stTcpLimitArea);
m_PassOnZones(vio_Visu := vio_Visu, vio_aZones := vo_Config.stActive.aZones, vi_un_Count := vo_Config.stActive.nZoneCount,
	vi_un_VisuCount := vio_Visu.vo_Visu.stConfig.nZoneCount);
m_PassOnFingers(vio_Visu := vio_Visu, vio_aFingers := vo_Config.stActive.aFingers,
	vi_un_Count := vo_Config.stActive.nFingerCount, vi_un_VisuCount := vio_Visu.vo_Visu.stConfig.nFingerCount);
END_METHOD

(****************************************************************************************************<br>
© Syntegon Group.<br>
All rights reserved, also regarding any disposal, exploitation, reproduction, editing, distribution,<br>
as well as in the event of applications for industrial property rights.<br>
*****************************************************************************************************<br>
DESCRIPTION:<br>
Effective pose of the track start (MCS), for the application's logic.<br>
****************************************************************************************************)
METHOD m_Pose : SynVisu.ST_VisuPose
m_Pose := vo_Config.stActive.stPose;
END_METHOD

END_FUNCTION_BLOCK

// ---- POUs/_FB_ConfigXtsLoop.TcPOU
(****************************************************************************************************<br>
© Syntegon Group.<br>
All rights reserved, also regarding any disposal, exploitation, reproduction, editing, distribution,<br>
as well as in the event of applications for industrial property rights.<br>
*****************************************************************************************************<br>
DESCRIPTION:<br>
Parameter set of one XTS loop (ADR 0017): its pose, origin shift, track modules, zones and gripper fingers,<br>
written by the configurator, taken over when the application allows it. Typical cycle:<br>
  fb_FxxParam.m_Register(vio_Manifest := GVL_Config.stManifest, vi_udn_Id := fb_Fxx.m_Id());<br>
  fb_FxxParam.m_Cycle(vio_Default := FxxDefault, vio_Set := FxxSet, vi_b_ApplyAllowed := b_Stopped);<br>
  fb_Fxx.m_Configure(vi_lr_ToolOffset := 120, ...);<br>
  fb_FxxParam.m_PassOn(vio_Visu := fb_Fxx);<br>
The application's logic takes its track and zones from m_Active, not from its own constants.<br>
*****************************************************************************************************<br>
OUTPUT VALUES:<br>
vo_Config is the contract structure the gateway reads and writes at the path in the config manifest.<br>
*****************************************************************************************************<br>
VERSION         ¦ DATE       ¦ NAME      ¦ CHANGE<br>
Syn_Config 1.1.0 ¦ 2026-11-10 ¦ J.Willner ¦ New<br>
Syn_Config 2.0.0 ¦ 2026-11-11 ¦ J.Willner ¦ Gripper fingers with their offsets (ADR 0018)<br>
Syn_Config 2.3.0 ¦ 2026-11-14 ¦ J.Willner ¦ m_Cycle through m_HandleStaging; m_PassOn passes the pose on<br>
****************************************************************************************************)
FUNCTION_BLOCK _FB_ConfigXtsLoop EXTENDS _FB_ConfigComponent
VAR_OUTPUT
	vo_Config							: ST_ConfigXtsLoop;	// contract structure of the gateway
END_VAR

(****************************************************************************************************<br>
© Syntegon Group.<br>
All rights reserved, also regarding any disposal, exploitation, reproduction, editing, distribution,<br>
as well as in the event of applications for industrial property rights.<br>
*****************************************************************************************************<br>
DESCRIPTION:<br>
All effective values (track modules, zones, ...), for the application's own logic.<br>
****************************************************************************************************)
METHOD m_Active : ST_ConfigXtsLoopParam
m_Active := vo_Config.stActive;
END_METHOD

(****************************************************************************************************<br>
© Syntegon Group.<br>
All rights reserved, also regarding any disposal, exploitation, reproduction, editing, distribution,<br>
as well as in the event of applications for industrial property rights.<br>
*****************************************************************************************************<br>
DESCRIPTION:<br>
An XTS loop.<br>
****************************************************************************************************)
METHOD PROTECTED m_ComponentType : SynVisu.E_VisuComponentType
m_ComponentType := SynVisu.E_VisuComponentType.XTS_LOOP;
END_METHOD

(****************************************************************************************************<br>
© Syntegon Group.<br>
All rights reserved, also regarding any disposal, exploitation, reproduction, editing, distribution,<br>
as well as in the event of applications for industrial property rights.<br>
*****************************************************************************************************<br>
DESCRIPTION:<br>
Every cycle: handles a staged set or a reset (a set only while vi_b_ApplyAllowed), keeps the active set in<br>
vio_Set and gives the effective values in vo_Config.stActive: the active set while one is valid, else the<br>
program values vio_Default.<br>
*****************************************************************************************************<br>
OUTPUT VALUES:<br>
TRUE in the cycle a set was taken over or reset.<br>
****************************************************************************************************)
METHOD m_Cycle : BOOL
VAR_IN_OUT CONSTANT
	vio_Default							: ST_ConfigXtsLoopParam;	// the application's program values
END_VAR
VAR_IN_OUT
	vio_Set								: ST_ConfigXtsLoopSet;	// the application's VAR PERSISTENT active set
END_VAR
VAR_INPUT
	vi_b_ApplyAllowed					: BOOL;	// [-] a staged set may be taken over now, e.g. while the machine stands
END_VAR
VAR
	b_TempTakeOver						: BOOL;	// the staged set was taken over: copy it
END_VAR
m_Cycle := m_HandleStaging(vio_Staging := vo_Config.stStaging, vio_Status := vo_Config.stStatus, vio_b_Valid := vio_Set.bValid,
	vio_udn_Version := vio_Set.nVersion, vio_udn_LastVersion := vio_Set.nLastVersion, vi_b_ApplyAllowed := vi_b_ApplyAllowed,
	vo_b_TakeOver => b_TempTakeOver);
IF b_TempTakeOver THEN
	vio_Set.stParam := vo_Config.stStaged;
END_IF


(****************************************************************************************************
EFFECTIVE VALUES
****************************************************************************************************)
IF vio_Set.bValid THEN
	vo_Config.stActive := vio_Set.stParam;
ELSE
	vo_Config.stActive := vio_Default;
END_IF
END_METHOD

(****************************************************************************************************<br>
© Syntegon Group.<br>
All rights reserved, also regarding any disposal, exploitation, reproduction, editing, distribution,<br>
as well as in the event of applications for industrial property rights.<br>
*****************************************************************************************************<br>
DESCRIPTION:<br>
Why a staged set cannot be taken over; '' when it can: a track without modules, more modules, zones or fingers<br>
than the lists hold, a module without a length, a zone on no conveyor (id 0), or a finger without a diameter or<br>
height.<br>
****************************************************************************************************)
METHOD PROTECTED m_InvalidStaged : STRING(80)
m_InvalidStaged := m_InvalidModules(vio_aModules := vo_Config.stStaged.aModules, vi_un_Count := vo_Config.stStaged.nModuleCount);
IF m_InvalidStaged = '' THEN
	m_InvalidStaged := m_InvalidZones(vio_aZones := vo_Config.stStaged.aZones, vi_un_Count := vo_Config.stStaged.nZoneCount);
END_IF
IF m_InvalidStaged = '' THEN
	m_InvalidStaged := m_InvalidFingers(vio_aFingers := vo_Config.stStaged.aFingers, vi_un_Count := vo_Config.stStaged.nFingerCount);
END_IF
END_METHOD

(****************************************************************************************************<br>
© Syntegon Group.<br>
All rights reserved, also regarding any disposal, exploitation, reproduction, editing, distribution,<br>
as well as in the event of applications for industrial property rights.<br>
*****************************************************************************************************<br>
DESCRIPTION:<br>
Passes the effective pose, origin shift, track modules, zones and fingers on to the loop's Syn_Visu FB, so the<br>
visualisation shows what the machine uses; the tool offset and mover size (hardware) stay with the<br>
application's m_Configure call. Call it after m_Cycle, every cycle; Syn_Visu's config version only changes when<br>
a value does.<br>
****************************************************************************************************)
METHOD m_PassOn : BOOL
VAR_IN_OUT
	vio_Visu							: SynVisu._FB_VisuXtsLoop;	// the loop's Syn_Visu FB
END_VAR
m_PassOn := TRUE;
vio_Visu.m_SetPose(vi_Pose := vo_Config.stActive.stPose);
vio_Visu.m_SetOriginShift(vi_lr_X := vo_Config.stActive.stOriginShift.fX, vi_lr_Y := vo_Config.stActive.stOriginShift.fY,
	vi_lr_Z := vo_Config.stActive.stOriginShift.fZ);
m_PassOnModules(vio_Visu := vio_Visu, vio_aModules := vo_Config.stActive.aModules,
	vi_un_Count := vo_Config.stActive.nModuleCount, vi_un_VisuCount := vio_Visu.vo_Visu.stConfig.nModuleCount);
m_PassOnZones(vio_Visu := vio_Visu, vio_aZones := vo_Config.stActive.aZones, vi_un_Count := vo_Config.stActive.nZoneCount,
	vi_un_VisuCount := vio_Visu.vo_Visu.stConfig.nZoneCount);
m_PassOnFingers(vio_Visu := vio_Visu, vio_aFingers := vo_Config.stActive.aFingers,
	vi_un_Count := vo_Config.stActive.nFingerCount, vi_un_VisuCount := vio_Visu.vo_Visu.stConfig.nFingerCount);
END_METHOD

(****************************************************************************************************<br>
© Syntegon Group.<br>
All rights reserved, also regarding any disposal, exploitation, reproduction, editing, distribution,<br>
as well as in the event of applications for industrial property rights.<br>
*****************************************************************************************************<br>
DESCRIPTION:<br>
Effective pose of the start of module 1 (MCS), for the application's logic.<br>
****************************************************************************************************)
METHOD m_Pose : SynVisu.ST_VisuPose
m_Pose := vo_Config.stActive.stPose;
END_METHOD

END_FUNCTION_BLOCK
